FUNCTION_BLOCK basicMotorInovaisa (* Status de um motor do painel do gradeamento (grade ou rosca) *)
  (* Standard: 61499-2 *)
  (* Version 1.0, 22/10/2026, Hidryco, Hidryco, 1.0: codigos de funcionamento da tabela Inovaisa PV-35524 (grade com reverso, rosca), sobretorque, falha *)
  PACKAGE Hidryco.HidrycoLib;
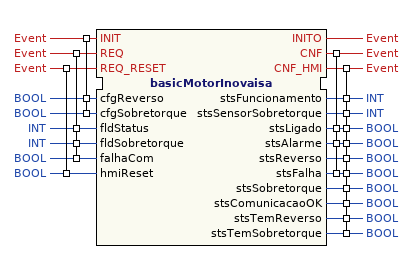
  EVENT_INPUT
    INIT WITH cfgReverso, cfgSobretorque; (* Inicializacao (configuracao da instancia) *)
    REQ WITH fldStatus, fldSobretorque, falhaCom; (* Leitura do painel (pelo processo) *)
    REQ_RESET WITH hmiReset; (* IHM: reconhece os alarmes *)
  END_EVENT
  EVENT_OUTPUT
    INITO; (* Inicializacao concluida *)
    CNF WITH stsLigado, stsFalha, stsAlarme; (* Status para o processo (na mudanca) *)
    CNF_HMI WITH stsFuncionamento, stsSensorSobretorque, stsLigado, stsAlarme, stsReverso, stsFalha, stsSobretorque, stsComunicacaoOK, stsTemReverso, stsTemSobretorque; (* Status para a IHM e alarmes (na mudanca) *)
  END_EVENT
  VAR_INPUT
    cfgReverso : BOOL := FALSE; (* TRUE = grade (codigos 0 parado, 1 avante, 2 reverso, 3 falha); FALSE = rosca (0 parado, 1 funcionando, 2 falha) *)
    cfgSobretorque : BOOL := FALSE; (* TRUE = tem sensor de sobretorque *)
    fldStatus : INT; (* Registro de status do motor (4007/4008/4009) *)
    fldSobretorque : INT; (* Registro do sobretorque (4010/4011) *)
    falhaCom : BOOL; (* Sem comunicacao com o painel *)
    hmiReset : BOOL; (* IHM: reconhece os alarmes *)
  END_VAR
  VAR_OUTPUT
    stsFuncionamento : INT; (* Codigo de funcionamento do painel: grade 0 parado, 1 avante, 2 reverso, 3 falha; rosca 0 parado, 1 funcionando, 2 falha *)
    stsSensorSobretorque : INT; (* Sensor de sobretorque: 0 normal, 1 sobretorque (so grade) *)
    stsLigado : BOOL; (* Motor funcionando (avante ou reverso) *)
    stsAlarme : BOOL; (* Falha do motor ou sobretorque *)
    stsReverso : BOOL; (* Grade funcionando em reverso *)
    stsFalha : BOOL; (* Motor em falha (informado pelo painel) *)
    stsSobretorque : BOOL; (* Sobretorque atuado *)
    stsComunicacaoOK : BOOL; (* Comunicacao com o painel do gradeamento OK *)
    stsTemReverso : BOOL; (* Configuracao: motor com reverso (grade) *)
    stsTemSobretorque : BOOL; (* Configuracao: motor com sensor de sobretorque (grade) *)
  END_VAR
  VAR
    initDone : BOOL;
    recebido : BOOL;
    primeiro : BOOL := TRUE;
    sig : INT;
    oldSig : INT := -1;
  END_VAR
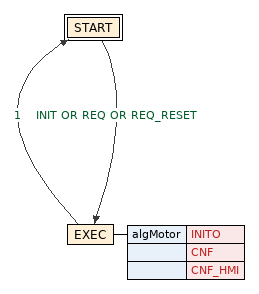
  EC_STATES
    START; (* Estado inicial *)
    EXEC : algMotor -> INITO, -> CNF, -> CNF_HMI; (* Executa a logica; o algoritmo decide quais eventos saem *)
  END_STATES
  EC_TRANSITIONS
    START TO EXEC := INIT OR REQ OR REQ_RESET;
    EXEC TO START := 1;
  END_TRANSITIONS
  ALGORITHM algMotor IN ST: (* Logica completa *)
(* =====================================================================
   basicMotorInovaisa v1.0 - status de um motor do painel do gradeamento
   (Vibropac PV-35524, tabela Modbus Inovaisa): o painel comanda o motor;
   aqui so a leitura do estado, a falha e o sobretorque (sem memoria:
   seguem o painel; o reconhecimento fica nos alarmes).
   ===================================================================== *)
INITO   := FALSE;
CNF     := FALSE;
CNF_HMI := FALSE;
IF INIT THEN
    initDone := TRUE;
    INITO := TRUE;
END_IF;
IF NOT initDone THEN
    RETURN;
END_IF;
IF REQ THEN
    recebido := TRUE;
END_IF;
stsTemReverso := cfgReverso;
stsTemSobretorque := cfgSobretorque;
stsComunicacaoOK := recebido AND NOT falhaCom;
IF stsComunicacaoOK THEN
    stsFuncionamento := fldStatus;
    IF cfgReverso THEN
        stsLigado  := (fldStatus = 1) OR (fldStatus = 2);
        stsReverso := fldStatus = 2;
        stsFalha   := fldStatus = 3;
    ELSE
        stsLigado  := fldStatus = 1;
        stsReverso := FALSE;
        stsFalha   := fldStatus = 2;
    END_IF;
    IF cfgSobretorque THEN
        stsSensorSobretorque := fldSobretorque;
    ELSE
        stsSensorSobretorque := 0;
    END_IF;
    stsSobretorque := cfgSobretorque AND (fldSobretorque <> 0);
ELSE
    stsFuncionamento := 0;
    stsSensorSobretorque := 0;
    stsLigado := FALSE;
    stsReverso := FALSE;
    stsFalha := FALSE;
    stsSobretorque := FALSE;
END_IF;
stsAlarme := stsFalha OR stsSobretorque;
sig := stsFuncionamento * 16 + stsSensorSobretorque;
IF stsComunicacaoOK THEN sig := sig + 4096; END_IF;
IF primeiro OR (sig <> oldSig) THEN
    CNF := TRUE;
    CNF_HMI := TRUE;
END_IF;
IF REQ_RESET THEN
    CNF_HMI := TRUE;
END_IF;
oldSig := sig;
primeiro := FALSE;
  END_ALGORITHM
END_FUNCTION_BLOCK
